(* PLC project v0.5.8_.project, CODESYS CODESYS V3.5 SP19 Patch 1 *)
(* stored: creationDateTime 2026-08-05T11:24:59.5567926, modificationDateTime 2026-08-05T05:05:15.4109854 *)

CONFIGURATION LocalDevice
END_CONFIGURATION

CONFIGURATION Local_Digital_IO
END_CONFIGURATION

CONFIGURATION EtherCAT_Master
END_CONFIGURATION

CONFIGURATION Sendix_F58x8_1
END_CONFIGURATION

CONFIGURATION COD1_CODEUR
END_CONFIGURATION

CONFIGURATION Slot_2
END_CONFIGURATION

CONFIGURATION AC600_ECAT_Drive
END_CONFIGURATION

CONFIGURATION Sendix_F58x8_2
END_CONFIGURATION

CONFIGURATION COD2_CODEUR
END_CONFIGURATION

CONFIGURATION Slot_2_1
END_CONFIGURATION

CONFIGURATION VH_ExtensionDevice
END_CONFIGURATION

CONFIGURATION VH_0808ETP
END_CONFIGURATION

CONFIGURATION VH_0800END
END_CONFIGURATION

CONFIGURATION VH_0008ER
END_CONFIGURATION

CONFIGURATION VH_0008ER_1
END_CONFIGURATION

CONFIGURATION CANbus
END_CONFIGURATION

CONFIGURATION CANopen_Manager
END_CONFIGURATION

CONFIGURATION JOY1_JOYSTICK_MCB560_CO4201A
END_CONFIGURATION
